Staubli VAL3: initMsg.pgx

program initMsg()
  local num i
begin
  for i=0 to size(sRobotMsg)-1
    sRobotMsg[i]=""
  endFor
end
